Fanuc KAREL source: ka00091.KL

-- PROVISIONAL review KL for V1013-1; original PC SHA256 eed720c61208fb0620d3ffbcfb0b1db1f18884563c41f9a171de9af387da044f
-- Incomplete behavior may be omitted. Consult companion uncertainty JSON. Do not deploy.
PROGRAM KA00091
%NOLOCKGROUP
-- UNRESOLVED_DECL SRC type=000199
-- UNRESOLVED_DECL DST type=000106
BEGIN
  -- UNRESOLVED_PC offsets 5-25; opcodes 49,7E,4A
  -- UNRESOLVED_PC offsets 30-34; opcodes 7F
END KA00091
